FUNCTION_BLOCK Empty_cotrol (* Basic Function Block Type *)
  (* Standard: 61499-2 *)
  (* Version 0.0, 10/19/2026, lizar, Schneider Electric, Template *)
  PACKAGE Main;
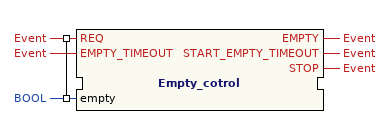
  EVENT_INPUT
    REQ WITH empty; (* Normal Execution Request *)
    EMPTY_TIMEOUT;
  END_EVENT
  EVENT_OUTPUT
    EMPTY;
    START_EMPTY_TIMEOUT;
    STOP;
  END_EVENT
  VAR_INPUT
    empty : BOOL; (* Input event qualifier *)
  END_VAR
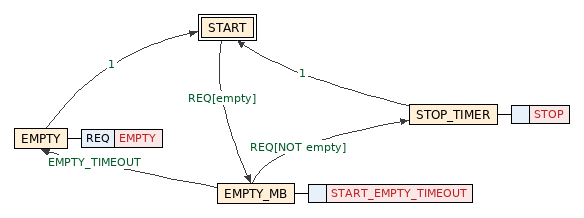
  EC_STATES
    START; (* Initial State *)
    EMPTY : REQ -> EMPTY; (* Normal execution *)
    EMPTY_MB : -> START_EMPTY_TIMEOUT;
    STOP_TIMER : -> STOP;
  END_STATES
  EC_TRANSITIONS
    START TO EMPTY_MB := REQ[empty];
    EMPTY_MB TO EMPTY := EMPTY_TIMEOUT;
    EMPTY_MB TO STOP_TIMER := REQ[NOT empty];
    EMPTY TO START := 1;
    STOP_TIMER TO START := 1;
  END_TRANSITIONS
  ALGORITHM REQ IN ST: (* Normally executed algorithm *)
;
  END_ALGORITHM
END_FUNCTION_BLOCK
